// TIA Portal V17 export
// export: Created 2026-11-08T05:50:31.5603516Z, ExportSetting WithDefaults, DisplayName Totally Integrated Automation Portal, DisplayVersion V17, DisplayName TIA Portal Openness, DisplayVersion V17, DisplayName TIA Portal Version Control Interface, DisplayVersion V17, DisplayName STEP 7 Professional, DisplayVersion V17, DisplayName STEP 7 Safety, DisplayVersion V17, DisplayName WinCC Professional, DisplayVersion V17
TagTable "HMI_Motor"
  Cmd_Marcha : Bool  (PLC tag DB_HMI.Cmd_Marcha, HMI_Connection_1, 100 ms)
  Cmd_Paro : Bool  (PLC tag DB_HMI.Cmd_Paro, HMI_Connection_1, 100 ms)
  Cmd_Reset : Bool  (PLC tag DB_HMI.Cmd_Reset, HMI_Connection_1, 100 ms)
  Sel_Estilo : Int  (PLC tag DB_HMI.Sel_Estilo, HMI_Connection_1, 100 ms)
  Estado : Int  (PLC tag DB_HMI.Estado, HMI_Connection_1, 100 ms)
  Motor_En_Marcha : Bool  (PLC tag DB_HMI.Motor_En_Marcha, HMI_Connection_1, 100 ms)
  Falla_Termico : Bool  (PLC tag DB_HMI.Falla_Termico, HMI_Connection_1, 100 ms)
  Pantalla : Int  (PLC tag DB_HMI.Pantalla, HMI_Connection_1, 100 ms)
  PB_Marcha : Bool  (PLC tag PB_Marcha, HMI_Connection_1, 100 ms)
  PB_Paro : Bool  (PLC tag PB_Paro, HMI_Connection_1, 100 ms)
  MOT1_Termico_Falla : Bool  (PLC tag MOT1_Termico_Falla, HMI_Connection_1, 100 ms)
  KM1_Motor : Bool  (PLC tag KM1_Motor, HMI_Connection_1, 100 ms)
  HL_Marcha : Bool  (PLC tag HL_Marcha, HMI_Connection_1, 100 ms)
  HL_Falla : Bool  (PLC tag HL_Falla, HMI_Connection_1, 100 ms)
  Banderas_Estado : Int  (PLC tag DB_Motor_Banderas.Estado, HMI_Connection_1, 100 ms)
  Banderas_Motor : Bool  (PLC tag DB_Motor_Banderas.Motor, HMI_Connection_1, 100 ms)
  Moore_Estado : Int  (PLC tag DB_Motor_Moore.Estado, HMI_Connection_1, 100 ms)
  Moore_Motor : Bool  (PLC tag DB_Motor_Moore.Motor, HMI_Connection_1, 100 ms)
  Mealy_Estado : Int  (PLC tag DB_Motor_Mealy.Estado, HMI_Connection_1, 100 ms)
  Mealy_Motor : Bool  (PLC tag DB_Motor_Mealy.Motor, HMI_Connection_1, 100 ms)
